TYPE "ST_CycleSummary"
VERSION : 0.1
   STRUCT
      CycleNo : UDInt;
      Started : LDT;
      StartedTimeSynchronized : Bool;
      Total : Time;
      WorkTime : Time;
      WaitTime : Time;
      ByClass : Array[0..4] of Time;
   END_STRUCT;

END_TYPE

